(* IEC 61131-3 sources: kns-port-domestic/targets/astra/src/POUs/Station/FB_StationAlarms, 6 files *)

(* ---- FB_StationAlarms.decl.st ---- *)
// Назначение: тревоги станции KNS1.* (04 §15, 05_alarm_list.csv) — 13 экземпляров PL.FB_Alarm,
//             индекс = E_StationAlarm, номер = STN_ALARM_ID_BASE + slot. Условия, подавления по
//             условию и значения задаёт PRG_Station; маски команд — бит slot - 1. Источник тревог
//             PL.I_AlarmSource для сводки (GetAlarm: индекс 0 — slot 1).
// Автор:      kr0nsch
// Версия:     0.1.0
// Документ:   docs/DESIGN.md, раздел 6.11; docs/04_algorithms.md, раздел 15
FUNCTION_BLOCK FB_StationAlarms IMPLEMENTS PL.I_AlarmSource
VAR_INPUT
    axCond       : ARRAY[1..GVL_Const.STN_ALARM_COUNT] OF BOOL;   // индекс — E_StationAlarm
    axSuppress   : ARRAY[1..GVL_Const.STN_ALARM_COUNT] OF BOOL;   // SuppressedByDesign
    arValue      : ARRAY[1..GVL_Const.STN_ALARM_COUNT] OF REAL;
    wAckReq      : WORD;            // маски stStationCmd, бит slot - 1
    wShelveReq   : WORD;
    wUnshelveReq : WORD;
    xAckAll      : BOOL;
    itfTime      : PL.I_TimeSource;
END_VAR
VAR_IN_OUT CONSTANT
    stCfg : ST_StationCfg;          // astAlarm[1..13]
END_VAR
VAR_OUTPUT
    wAlmActive  : WORD;
    wAlmUnack   : WORD;
    wAlmShelved : WORD;
    ePrioUnack  : PL.E_AlarmPriority;
END_VAR
VAR
    afbAlarm : ARRAY[1..GVL_Const.STN_ALARM_COUNT] OF PL.FB_Alarm;   // udiId = STN_ALARM_ID_BASE + slot
END_VAR
VAR_TEMP
    uiSlot : UINT;                  // слот тревоги
    wBit   : WORD;                  // бит слота в словах: slot - 1
    eState : PL.E_AlarmState;       // состояние тревоги после вызова
END_VAR

(* ---- AckAll.method.decl.st ---- *)
// Запрос «квитировать все тревоги станции»; выполняет ближайший вызов тела. TRUE — было что квитировать
METHOD PUBLIC AckAll : BOOL
VAR
    uiIdx : UINT;                   // слот тревоги
END_VAR

(* ---- AckAll.method.impl.st ---- *)
AckAll := FALSE;
FOR uiIdx := 1 TO GVL_Const.STN_ALARM_COUNT DO
    IF afbAlarm[uiIdx].Ack() THEN
        AckAll := TRUE;
    END_IF
END_FOR

(* ---- FB_StationAlarms.impl.st ---- *)
wAlmActive := 0;
wAlmUnack := 0;
wAlmShelved := 0;
ePrioUnack := PL.E_AlarmPriority.None;
FOR uiSlot := 1 TO GVL_Const.STN_ALARM_COUNT DO
    wBit := SHL(WORD#1, uiSlot - 1);
    // Запросы команд — до вызова тела: его выполняет вызов в этом же цикле (R3 контракта).
    // Shelve(T#0S) — на tShelveMax тревоги; при tShelveMax = 0 (EHL) FB_Alarm отклоняет запрос
    IF xAckAll OR (wAckReq AND wBit) <> 0 THEN
        afbAlarm[uiSlot].Ack();
    END_IF
    IF (wShelveReq AND wBit) <> 0 THEN
        afbAlarm[uiSlot].Shelve(tDuration := T#0S);
    END_IF
    IF (wUnshelveReq AND wBit) <> 0 THEN
        afbAlarm[uiSlot].Unshelve();
    END_IF
    // условие при подавлении не копит выдержку: после снятия подавления она отсчитывается заново. Иначе условие,
    // которое держится ещё цикл (станция видит выходы устройств циклом позже: после «сухого хода» и восстановления
    // питания насосы ещё «недоступны»), давало мелькание KNS1.NORES (High, сирена) — прогон ПМИ 19.10.2026
    afbAlarm[uiSlot](xIn := axCond[uiSlot] AND NOT axSuppress[uiSlot], xSuppress := axSuppress[uiSlot],
                     xOutOfService := FALSE,
                     udiId := GVL_Const.STN_ALARM_ID_BASE + UINT_TO_UDINT(uiSlot), rValue := arValue[uiSlot],
                     stCfg := stCfg.astAlarm[uiSlot], itfTime := itfTime);
    eState := afbAlarm[uiSlot].eState;
    IF afbAlarm[uiSlot].xActive THEN
        wAlmActive := wAlmActive OR wBit;
    END_IF
    IF afbAlarm[uiSlot].xUnacked THEN
        wAlmUnack := wAlmUnack OR wBit;
        IF TO_INT(afbAlarm[uiSlot].AlarmPriority) > TO_INT(ePrioUnack) THEN
            ePrioUnack := afbAlarm[uiSlot].AlarmPriority;
        END_IF
    END_IF
    // дополнение к активным: отложены оператором, подавлены логикой, выведены из работы
    IF eState = PL.E_AlarmState.Shelved OR eState = PL.E_AlarmState.SuppressedByDesign
       OR eState = PL.E_AlarmState.OutOfService THEN
        wAlmShelved := wAlmShelved OR wBit;
    END_IF
END_FOR

(* ---- GetAlarm.method.decl.st ---- *)
// Тревога по индексу источника: 0 — slot 1 (EHL) … STN_ALARM_COUNT - 1 — slot 13 (SIM); вне — 0
METHOD PUBLIC GetAlarm : PL.I_Alarm
VAR_INPUT
    uiIndex : UINT;                 // индекс 0…AlarmCount - 1
END_VAR

(* ---- GetAlarm.method.impl.st ---- *)
IF uiIndex < GVL_Const.STN_ALARM_COUNT THEN
    GetAlarm := afbAlarm[uiIndex + 1];
ELSE
    GetAlarm := 0;
END_IF
